{attribute 'qualified_only'}
{attribute 'strict'}
{attribute 'to_string'}
TYPE E_ASense_Name :
(
	eNotSelected := 0,
	//level sensors CIP	
	LT1004,	
	LT1003,	
	LT1002,
	LT1001,
	//Flow  sensors
	FT1001,
	FT1002,

	
	
	//conductivity sensors
	CT1101,
	CT3101,//not exist	
		
	//temperature sensors
	TT1001,
	TT1002,
	TT1003,
	TT1004,
	TT1101,
	TT1105,
	CT1101_2,
	CT1101_3,
	CT1101_4,
	TT2001,
	TT3001,
	TT3002,
	TT4001,
	TT4002,
	
	//level sensors


	LT1061,
	LT1071,
	LT3001,
	LT3002,
	LT4001,
	LT4002,
	
	//Pressure sensors
	PT1001,
	PT3001,
	PT3002,
	PT4001,
	PT4002,
	PT9001,
	PT9002,
	PT9011,

	FT4001,
	FT4002,	
	FT9011,
	
	//Air Pressure
	AP1001, //CIP
	AP2001, // TriBlender
	AP3001, //Marinade
	AP4001, //Color
	
	CT4101,	
	CT4102,	

	FT9012,
	
	//virtual list
	last
);
END_TYPE

(* stored: Version 1.1.0.1, ProductVersion 3.1.4024.13
   EnumerationTextList E_ASense_Name: Id {58e6c96c-1337-4953-b9cd-57c742ebe203} *)
